Fanuc KAREL source: KA00009.KL

PROGRAM KA00009
%NOLOCKGROUP
VAR
  SRC: INTEGER
  DST: VECTOR
BEGIN
  SRC = 2
  DST = SRC
END KA00009
